(* CODESYS project GVL_MAGAZINE_AXIS.gvl.xml

Project tree, tasks and I/O mapping:
  global variables GVL_MAGAZINE_AXIS
*)

// GVL_MAGAZINE_AXIS
{attribute 'qualified_only'}
VAR_GLOBAL
	// Legacy-объявление оставлено до удаления SoftMotion-узлов Magazine_1/2 через
	// CODESYS. Активная программа массив не читает, не пишет и FB_AXIS для него не создаёт.
	astAxis : ARRAY [1..GVL_CELL_SETTINGS.MagazineCount] OF ST_AXIS;
END_VAR
